TYPE "ST_ShiftRowV3"
VERSION : 0.1
   STRUCT
      StartMin : DInt := -1;
      DurationMin : DInt := 1440;
      ActiveDays : DInt;
      ProductionTarget : DInt;
   END_STRUCT;

END_TYPE

